(* IEC 61131-3 sources: Gen-AI/docs/member2_validation/codesys_release_v1.1/C03_syntax, 1 file *)

(* ---- source.st ---- *)
FUNCTION_BLOCK FB_AgentProbeSyntax
VAR_INPUT
 x : BOOL;
END_VAR
VAR_OUTPUT
 y : BOOL;
END_VAR
IF x y := TRUE; END_IF;
END_FUNCTION_BLOCK
